(* IEC 61131-3 sources: SemaPLC/sema-plc-benchmark/spec2control-benchmark/data/st-baseline/waste_water_treatment_facility/pous/programs, 8 files *)

(* ---- main.st ---- *)
PROGRAM main
VAR
	Heartbeat : bool;
END_VAR

(* Entry point required by OpenPLC Editor v4. The process sections run as parallel program instances under task0; main only provides a scan heartbeat. *)
Heartbeat := NOT Heartbeat;

END_PROGRAM

(* ---- Section10.st ---- *)
PROGRAM Section10
VAR
	FT_901_FlowRate : real;
	LS_901_LevelPercent : real;
	P_901A_Running : bool;
	P_901B_Running : bool;
	P_901AB_DutyActiveIsA : bool;
	P_901AB_SwitchedDueToDuty : bool;
	P_901AB_SwitchedDueToFailure : bool;
	FT_901 : ANALOG_IN;
	LS_901 : ANALOG_IN;
	P_901A : MOTOR_ON_OFF;
	P_901B : MOTOR_ON_OFF;
	XV_102 : VALVE_ON_OFF;
	P_901AB : DUTY_STANDBY;
	DutyTimer_TON : TON;
	FailA_TON : TON;
	FailB_TON : TON;
	SwitchoverDelay_TON : TON;
	AnyRunning_OR : bool;
	StartBand_AND : bool;
	LevelAbove60_GT : bool;
	LevelAbove40_GT : bool;
	LevelAbove85_GT : bool;
	StartRequest_OR : bool;
	FlowLessThan15_GT : bool;
	FailCondA_AND : bool;
	FailCondB_AND : bool;
	Failure_OR : bool;
	StartCmdA_OR : bool;
	StartCmdB_OR : bool;
	PumpA_Inhibit_OR : bool;
	PumpB_Inhibit_OR : bool;
	BothPumpsFailed_AND : bool;
END_VAR

FT_901(
    Alarm_Enable := TRUE);
LS_901(
    PV_High := 90.0,
    Alarm_Enable := TRUE);
FlowLessThan15_GT := (REAL#15.0 > FT_901.PV);
FailCondA_AND := P_901A.FB_Running AND FlowLessThan15_GT;
FailA_TON(
    IN := FailCondA_AND,
    PT := T#10s);
PumpA_Inhibit_OR := LS_901.Low_Alarm OR FailA_TON.Q OR P_901A.FB_Trip;
LevelAbove85_GT := (LS_901.PV > REAL#85.0);
FailCondB_AND := P_901B.FB_Running AND FlowLessThan15_GT;
FailB_TON(
    IN := FailCondB_AND,
    PT := T#10s);
PumpB_Inhibit_OR := LS_901.Low_Alarm OR FailB_TON.Q OR P_901B.FB_Trip;
StartCmdB_OR := LevelAbove85_GT OR P_901AB.CmdPumpB;
P_901B(
    Start_Cmd := StartCmdB_OR,
    MinRunTime := T#30m,
    Inhibit := PumpB_Inhibit_OR);
AnyRunning_OR := P_901A.FB_Running OR P_901B.FB_Running;
DutyTimer_TON(
    IN := AnyRunning_OR,
    PT := T#48h);
LevelAbove60_GT := (LS_901.PV > REAL#60.0);
LevelAbove40_GT := (LS_901.PV > REAL#40.0);
StartBand_AND := AnyRunning_OR AND LevelAbove40_GT;
StartRequest_OR := LevelAbove60_GT OR StartBand_AND;
Failure_OR := FailA_TON.Q OR FailB_TON.Q;
SwitchoverDelay_TON(
    IN := Failure_OR,
    PT := T#5s);
P_901AB(
    Enable := TRUE,
    StartRequest := StartRequest_OR,
    AlternateEnable := TRUE,
    DutyElapsed := DutyTimer_TON.Q,
    SwitchoverDelayElapsed := SwitchoverDelay_TON.Q,
    PumpA_RunFB := P_901A.FB_Running,
    PumpB_RunFB := P_901B.FB_Running,
    PumpA_Fault := FailA_TON.Q,
    PumpB_Fault := FailB_TON.Q);
StartCmdA_OR := LevelAbove85_GT OR P_901AB.CmdPumpA;
P_901A(
    Start_Cmd := StartCmdA_OR,
    MinRunTime := T#30m,
    Inhibit := PumpA_Inhibit_OR);
BothPumpsFailed_AND := FailA_TON.Q AND FailB_TON.Q;
XV_102(
    Inhibit := BothPumpsFailed_AND);

(* Outputs published to other sections / HMI. *)
FT_901_FlowRate := FT_901.PV;
LS_901_LevelPercent := LS_901.PV;
P_901A_Running := P_901A.FB_Running;
P_901B_Running := P_901B.FB_Running;
P_901AB_DutyActiveIsA := P_901AB.ActiveIsA;
P_901AB_SwitchedDueToDuty := P_901AB.SwitchedDueToDuty;
P_901AB_SwitchedDueToFailure := P_901AB.SwitchedDueToFailure;

END_PROGRAM

(* ---- Section11.st ---- *)
PROGRAM Section11
VAR
	FIT_104_InfluentFlow_PV : real;
	FIC_106_SP_From_FFIC_107 : real;
	FIT_104 : ANALOG_IN;
	FFIC_107 : RATIO_CONTROL;
	FIC_106 : PID_BASIC;
	CD_1001 : MOTOR_VSD;
	PV_101 : VALVE_ELECTRIC;
	XV_102 : VALVE_ON_OFF;
	PumpInhibitAggregator : bool;
	RatioCtrlInhibitAggregator : bool;
	PumpOpenedInverter : bool;
END_VAR

FIT_104(
    Scaling_Slope := 6.25,
    Scaling_Offset := -25.0,
    Alarm_Enable := TRUE);
FIC_106(
    AUTO := TRUE,
    PV := CD_1001.FB_ActualSpeed,
    SP := FFIC_107.SlaveSP,
    MV_MIN := 0.0,
    MV_MAX := 100.0,
    Deviation_Limit := 3.0);
PV_101(
    Open_Limit := 100.0,
    Close_Limit := 0.0);
XV_102();
PumpOpenedInverter := NOT XV_102.FB_Opened;
PumpInhibitAggregator := PumpOpenedInverter OR FIT_104.Low_Alarm OR FIT_104.General_Fault OR XV_102.Alarm_General OR XV_102.Alarm_Position_Error OR PV_101.Alarm OR PV_101.Position_Error OR CD_1001.Alarm_Comm_Fail OR CD_1001.FB_Fault OR CD_1001.Alarm_Speed_Deviation;
CD_1001(
    Speed_SP := FIC_106.XOUT,
    Inhibit := PumpInhibitAggregator);
RatioCtrlInhibitAggregator := FIT_104.Low_Alarm OR FIT_104.High_Alarm OR FIT_104.General_Fault OR CD_1001.FB_Fault OR CD_1001.Alarm_Comm_Fail OR CD_1001.Alarm_Speed_Deviation;
FFIC_107(
    Auto := TRUE,
    PrimaryPV := FIT_104.PV,
    SecondaryPV := CD_1001.FB_ActualSpeed,
    RatioSP := 2.5,
    Bias := 0.0,
    MV_MIN := 0.0,
    MV_MAX := 100.0,
    Inhibit := RatioCtrlInhibitAggregator);

(* Outputs published to other sections / HMI. *)
FIT_104_InfluentFlow_PV := FIT_104.PV;
FIC_106_SP_From_FFIC_107 := FFIC_107.SlaveSP;

END_PROGRAM

(* ---- Section12.st ---- *)
PROGRAM Section12
VAR
	IIC101_Raw_mA : real;
	LV104_Raw_mA : real;
	IIC101_Solids_PV : real;
	IIC103_MV_to_PV102 : real;
	LV104_Level_PV : real;
	IIC_101 : ANALOG_IN;
	LV_104 : ANALOG_IN;
	IIC_103 : PID_BASIC;
	IIC_105 : BOOL_INPUT;
	PV_102 : VALVE_ELECTRIC;
	OC_1101 : VALVE_ON_OFF;
	OdorNotActive_NOT : bool;
	PIDInhibit_OR : bool;
	ValveInhibit_OR : bool;
END_VAR

IIC_101(
    Raw_Signal := IIC101_Raw_mA,
    Scaling_Slope := 0.625,
    Scaling_Offset := -2.5,
    Alarm_Enable := TRUE);
LV_104(
    Raw_Signal := LV104_Raw_mA,
    PV_High := 85.0,
    Scaling_Slope := 6.25,
    Scaling_Offset := -25.0,
    Alarm_Enable := TRUE);
PIDInhibit_OR := LV_104.High_Alarm OR IIC_101.General_Fault;
OC_1101(
    Timeout := T#10s);
IIC_105(
    Bool_In := OC_1101.FB_Opened);
OdorNotActive_NOT := NOT IIC_105.Bool_Out;
ValveInhibit_OR := OdorNotActive_NOT OR PV_102.Position_Error;
PV_102(
    Control_Signal := IIC_103.XOUT,
    Manual_Mode := FALSE,
    Open_Limit := 100.0,
    Close_Limit := 0.0,
    Timeout := T#30s,
    Inhibit := ValveInhibit_OR);
IIC_103(
    AUTO := TRUE,
    PV := IIC_101.PV,
    SP := 6.5,
    MV_MIN := 10.0,
    MV_MAX := 90.0,
    X0 := PV_102.Feedback_Pos,
    KP := 3.0,
    TR := 1.2,
    TD := 0.3,
    PV_High := 8.0,
    PV_Low := 4.0,
    Inhibit := PIDInhibit_OR);

(* Outputs published to other sections / HMI. *)
IIC101_Solids_PV := IIC_101.PV;
IIC103_MV_to_PV102 := IIC_103.XOUT;
LV104_Level_PV := LV_104.PV;

END_PROGRAM

(* ---- Section2.st ---- *)
PROGRAM Section2
VAR
	LS_101_WetWellLevel_PV_m : real;
	FT_101_InfluentFlow_PV_m3ph : real;
	PIC_101_WetWellLevel_MV_Pct : real;
	P_101A_Speed_Command_Pct : real;
	P_101B_Speed_Command_Pct : real;
	P101_LevelTrips_Active : bool;
	VG101_Inhibit_Active : bool;
	BS101_Disable_Active : bool;
	P_101A_Start_Cmd : bool;
	P_101B_Start_Cmd : bool;
	FT_101 : ANALOG_IN;
	LS_101 : ANALOG_IN;
	PIC_101 : PID_BASIC;
	P_101A : MOTOR_VSD;
	P_101B : MOTOR_VSD;
	XV_101 : VALVE_ON_OFF;
	BS_101 : BOOL_INPUT;
	VG_101 : MOTOR_ON_OFF;
	P101_LevelTrips_OR : bool;
	VG101_Inhibit_OR : bool;
	BS101_Disable_OR : bool;
	PID_Output_Positive_GT : bool;
	P101_LevelTrips_NOT : bool;
	PumpRunEnable_AND : bool;
	StartA_NOT : bool;
	StartB_NOT : bool;
	P101A_Running_NOT : bool;
	P101A_Failure_OR : bool;
	P101B_Start_AND : bool;
	LS101_HighAlarm_NOT : bool;
END_VAR

FT_101(
    Scaling_Slope := 31.25,
    Scaling_Offset := -125.0,
    Alarm_Enable := TRUE);
LS_101(
    PV_High := 8.5,
    PV_Low := 1.5,
    Scaling_Slope := 0.625,
    Scaling_Offset := -2.5,
    Alarm_Enable := TRUE);
PIC_101(
    AUTO := TRUE,
    PV := LS_101.PV,
    SP := 5.5,
    MV_MIN := 30.0,
    MV_MAX := 90.0,
    X0 := 0.0,
    KP := -2.0,
    TR := 1.5,
    TD := 0.3,
    Deviation_Limit := 0.1);
P101_LevelTrips_OR := PIC_101.PV_Low_Alarm OR PIC_101.PV_High_Alarm OR LS_101.High_Alarm;
P101_LevelTrips_NOT := NOT P101_LevelTrips_OR;
PumpRunEnable_AND := P101_LevelTrips_NOT;
StartA_NOT := NOT PumpRunEnable_AND;
P_101A(
    Start_Cmd := PumpRunEnable_AND,
    Stop_Cmd := StartA_NOT,
    Speed_SP := PIC_101.XOUT,
    Inhibit := P101_LevelTrips_OR);
P101A_Running_NOT := NOT P_101A.FB_Running;
P101A_Failure_OR := P_101A.FB_Fault OR P101A_Running_NOT;
P101B_Start_AND := PumpRunEnable_AND AND P101A_Failure_OR;
StartB_NOT := NOT P101B_Start_AND;
P_101B(
    Start_Cmd := P101B_Start_AND,
    Stop_Cmd := StartB_NOT,
    Speed_SP := PIC_101.XOUT,
    Inhibit := P101_LevelTrips_OR);
LS101_HighAlarm_NOT := NOT LS_101.High_Alarm;
XV_101(
    Open_Cmd := LS101_HighAlarm_NOT,
    Close_Cmd := LS_101.High_Alarm);
BS101_Disable_OR := PIC_101.PV_Low_Alarm OR LS_101.Low_Alarm;
BS_101(
    Bool_In := BS101_Disable_OR);
VG101_Inhibit_OR := LS_101.Low_Alarm OR FT_101.Low_Alarm;
VG_101(
    Inhibit := VG101_Inhibit_OR);
PID_Output_Positive_GT := (0.0 > 0.0);

(* Outputs published to other sections / HMI. *)
P101_LevelTrips_Active := P101_LevelTrips_OR;
VG101_Inhibit_Active := VG101_Inhibit_OR;
BS101_Disable_Active := BS101_Disable_OR;
P_101A_Start_Cmd := PumpRunEnable_AND;
P_101B_Start_Cmd := P101B_Start_AND;
LS_101_WetWellLevel_PV_m := LS_101.PV;
FT_101_InfluentFlow_PV_m3ph := FT_101.PV;
PIC_101_WetWellLevel_MV_Pct := PIC_101.XOUT;
P_101A_Speed_Command_Pct := P_101A.Speed_Out;
P_101B_Speed_Command_Pct := P_101B.Speed_Out;

END_PROGRAM

(* ---- Section4.st ---- *)
PROGRAM Section4
VAR
	FT301_InfluentFlow_PV : real;
	FT302_SludgeFlow_PV : real;
	LS301_WeirLevel_PV : real;
	PS301_SludgePressure_PV : real;
	FT302_SludgeFlow_SP : real;
	FT_301 : ANALOG_IN;
	FT_302 : ANALOG_IN;
	LS_301 : ANALOG_IN;
	PS_301 : ANALOG_IN;
	SS_301 : DIGITAL_IN;
	FV_102 : VALVE_ELECTRIC;
	FFIC_303 : RATIO_CONTROL;
	FIC_302 : PID_BASIC;
	FlowAboveCutoff_GT : bool;
	MasterInhibit_OR : bool;
END_VAR

FT_301(
    Alarm_Enable := TRUE);
FT_302(
    Alarm_Enable := TRUE);
LS_301(
    PV_High := 5.0,
    PV_Low := 2.0,
    Alarm_Enable := TRUE);
PS_301();
SS_301();
FlowAboveCutoff_GT := (FT_301.PV > 50.0);
MasterInhibit_OR := LS_301.High_Alarm OR LS_301.Low_Alarm OR FT_301.High_Alarm OR FT_301.Low_Alarm OR FT_301.General_Fault OR FT_302.High_Alarm OR FT_302.Low_Alarm OR FT_302.General_Fault OR FIC_302.Deviation_Alarm OR FV_102.Position_Error OR FV_102.Alarm OR SS_301.DI_Out;
FFIC_303(
    Auto := FlowAboveCutoff_GT,
    PrimaryPV := FT_301.PV,
    SecondaryPV := FT_302.PV,
    RatioSP := 0.3,
    Bias := 0.0,
    TrimKp := 0.0,
    TrimTi := T#0s,
    MV_MIN := 0.0,
    MV_MAX := 200.0,
    Inhibit := MasterInhibit_OR);
FIC_302(
    AUTO := FlowAboveCutoff_GT,
    PV := FT_302.PV,
    SP := FFIC_303.SlaveSP,
    MV_MIN := 0.0,
    MV_MAX := 100.0,
    Deviation_Limit := 10.0,
    Inhibit := MasterInhibit_OR);
FV_102(
    Control_Signal := FIC_302.XOUT,
    Manual_Mode := MasterInhibit_OR,
    Manual_Position := 0.0,
    Inhibit := MasterInhibit_OR);

(* Outputs published to other sections / HMI. *)
FT301_InfluentFlow_PV := FT_301.PV;
FT302_SludgeFlow_PV := FT_302.PV;
LS301_WeirLevel_PV := LS_301.PV;
PS301_SludgePressure_PV := PS_301.PV;
FT302_SludgeFlow_SP := FFIC_303.SlaveSP;

END_PROGRAM

(* ---- Section7.st ---- *)
PROGRAM Section7
VAR
	PT_601A_DischargePressure_PV : real;
	PT_601B_DischargePressure_PV : real;
	CL_601_ActiveIsA : bool;
	PS_601_ActiveIsA : bool;
	CL_601A : MOTOR_ON_OFF;
	CL_601B : MOTOR_ON_OFF;
	PS_601A : MOTOR_ON_OFF;
	PS_601B : MOTOR_ON_OFF;
	PT_601A : ANALOG_IN;
	PT_601B : ANALOG_IN;
	LS_601 : DIGITAL_IN;
	VS_601A : VALVE_ELECTRIC;
	VS_601B : VALVE_ELECTRIC;
	CL_601A_CL_601B : DUTY_STANDBY;
	PS_601A_PS_601B : DUTY_STANDBY;
	Clar_MinRunTimer_TON : TON;
	Clar_DutyTimer_TON : TON;
	Clar_SwitchoverDelay_TON : TON;
	Pump_MinRunTimer_TON : TON;
	Pump_DutyTimer_TON : TON;
	Pump_SwitchoverDelay_TON : TON;
	ClarifierAnyRunning_OR : bool;
	ClarifierNoneRunning_NOT : bool;
	PumpAnyRunning_OR : bool;
	PumpNoneRunning_NOT : bool;
	PS601A_Inhibit_OR : bool;
	PS601B_Inhibit_OR : bool;
END_VAR

LS_601();
CL_601B(
    Start_Cmd := CL_601A_CL_601B.CmdPumpB,
    Start_Delay := T#5s,
    MinRunTime := T#30m,
    Inhibit := LS_601.DI_Out);
ClarifierAnyRunning_OR := CL_601A.FB_Running OR CL_601B.FB_Running;
Clar_DutyTimer_TON(
    IN := ClarifierAnyRunning_OR,
    PT := T#72h);
Clar_MinRunTimer_TON(
    IN := ClarifierAnyRunning_OR,
    PT := T#30m);
ClarifierNoneRunning_NOT := NOT ClarifierAnyRunning_OR;
Clar_SwitchoverDelay_TON(
    IN := ClarifierNoneRunning_NOT,
    PT := T#10s);
CL_601A_CL_601B(
    Enable := TRUE,
    StartRequest := TRUE,
    AlternateEnable := TRUE,
    DutyElapsed := Clar_DutyTimer_TON.Q,
    MinRunElapsed := Clar_MinRunTimer_TON.Q,
    SwitchoverDelayElapsed := Clar_SwitchoverDelay_TON.Q,
    PumpA_RunFB := CL_601A.FB_Running,
    PumpB_RunFB := CL_601B.FB_Running,
    PumpA_Fault := CL_601A.FB_Trip,
    PumpB_Fault := CL_601B.FB_Trip,
    Inhibit := LS_601.DI_Out);
CL_601A(
    Start_Cmd := CL_601A_CL_601B.CmdPumpA,
    Start_Delay := T#5s,
    MinRunTime := T#30m,
    Inhibit := LS_601.DI_Out);
PT_601A(
    PV_Low := 25.0,
    Alarm_Enable := TRUE);
PS601A_Inhibit_OR := PT_601A.Low_Alarm OR LS_601.DI_Out;
PT_601B(
    PV_Low := 25.0,
    Alarm_Enable := TRUE);
PS601B_Inhibit_OR := PT_601B.Low_Alarm OR LS_601.DI_Out;
PS_601B(
    Start_Cmd := PS_601A_PS_601B.CmdPumpB,
    Start_Delay := T#5s,
    MinRunTime := T#30m,
    Inhibit := PS601B_Inhibit_OR);
PumpAnyRunning_OR := PS_601A.FB_Running OR PS_601B.FB_Running;
Pump_DutyTimer_TON(
    IN := PumpAnyRunning_OR,
    PT := T#72h);
Pump_MinRunTimer_TON(
    IN := PumpAnyRunning_OR,
    PT := T#30m);
PumpNoneRunning_NOT := NOT PumpAnyRunning_OR;
Pump_SwitchoverDelay_TON(
    IN := PumpNoneRunning_NOT,
    PT := T#10s);
PS_601A_PS_601B(
    Enable := TRUE,
    StartRequest := TRUE,
    AlternateEnable := TRUE,
    DutyElapsed := Pump_DutyTimer_TON.Q,
    MinRunElapsed := Pump_MinRunTimer_TON.Q,
    SwitchoverDelayElapsed := Pump_SwitchoverDelay_TON.Q,
    PumpA_RunFB := PS_601A.FB_Running,
    PumpB_RunFB := PS_601B.FB_Running,
    PumpA_Fault := PS_601A.FB_Trip,
    PumpB_Fault := PS_601B.FB_Trip,
    Inhibit := LS_601.DI_Out);
PS_601A(
    Start_Cmd := PS_601A_PS_601B.CmdPumpA,
    Start_Delay := T#5s,
    MinRunTime := T#30m,
    Inhibit := PS601A_Inhibit_OR);
VS_601A(
    Open_Limit := 100.0,
    Close_Limit := 0.0);
VS_601B(
    Open_Limit := 100.0,
    Close_Limit := 0.0);

(* Outputs published to other sections / HMI. *)
PT_601A_DischargePressure_PV := PT_601A.PV;
PT_601B_DischargePressure_PV := PT_601B.PV;
CL_601_ActiveIsA := CL_601A_CL_601B.ActiveIsA;
PS_601_ActiveIsA := PS_601A_PS_601B.ActiveIsA;

END_PROGRAM

(* ---- Section9.st ---- *)
PROGRAM Section9
VAR
	FT_801_EffluentFlow_PV : real;
	CL_801_ChlorineFlow_SP : real;
	DC_801_DechlorFlow_SP : real;
	XV_106_FullyOpen_FB : bool;
	CL_801_Running_FB : bool;
	DC_801_Running_FB : bool;
	FT_801 : ANALOG_IN;
	FIC_101 : RATIO_CONTROL;
	FIC_102 : RATIO_CONTROL;
	CL_801 : MOTOR_VSD;
	DC_801 : MOTOR_VSD;
	LV_105 : VALVE_ELECTRIC;
	XV_106 : VALVE_ON_OFF;
	UV_801 : MOTOR_ON_OFF;
	CL_RatioMinCalc : real;
	CL_RatioMaxCalc : real;
	DC_RatioMinCalc : real;
	DC_RatioMaxCalc : real;
	ValveNotOpen : bool;
	CL_NotRunning : bool;
	ChemActive : bool;
	LV_105_AnyAlarm : bool;
	XV_106_AnyAlarm : bool;
	CL_801_Inh_OR1 : bool;
	CL_801_Inh_OR2 : bool;
	CL_801_Inh_OR3 : bool;
	DC_801_Inh_OR1 : bool;
	DC_801_Inh_OR2 : bool;
	FT_801_AnyFault_OR1 : bool;
	FT_801_AnyFault_OR2 : bool;
	FIC_102_Inh_OR1 : bool;
END_VAR

FT_801(
    Scaling_Slope := 62.5,
    Scaling_Offset := -250.0,
    Alarm_Enable := TRUE);
XV_106(
    Timeout := T#5s);
ValveNotOpen := NOT XV_106.FB_Opened;
CL_801_Inh_OR1 := ValveNotOpen OR FT_801.Low_Alarm;
XV_106_AnyAlarm := XV_106.Alarm_Position_Error OR XV_106.Alarm_General;
CL_801_Inh_OR2 := CL_801_Inh_OR1 OR XV_106_AnyAlarm;
LV_105(
    Timeout := T#5s);
LV_105_AnyAlarm := LV_105.Position_Error OR LV_105.Alarm;
CL_801_Inh_OR3 := CL_801_Inh_OR2 OR LV_105_AnyAlarm;
CL_801(
    Speed_SP := FIC_101.SlaveSP,
    Inhibit := CL_801_Inh_OR3);
CL_RatioMaxCalc := FT_801.PV * 3.0;
CL_RatioMinCalc := FT_801.PV * 2.0;
FT_801_AnyFault_OR1 := FT_801.Low_Alarm OR FT_801.High_Alarm;
FT_801_AnyFault_OR2 := FT_801_AnyFault_OR1 OR FT_801.General_Fault;
FIC_101(
    Auto := TRUE,
    PrimaryPV := FT_801.PV,
    SecondaryPV := CL_801.FB_ActualSpeed,
    RatioSP := 2.5,
    MV_MIN := CL_RatioMinCalc,
    MV_MAX := CL_RatioMaxCalc,
    Inhibit := FT_801_AnyFault_OR2);
CL_NotRunning := NOT CL_801.FB_Running;
DC_801_Inh_OR1 := LV_105_AnyAlarm OR FT_801.Low_Alarm;
DC_801_Inh_OR2 := DC_801_Inh_OR1 OR CL_NotRunning;
DC_801(
    Speed_SP := FIC_102.SlaveSP,
    Inhibit := DC_801_Inh_OR2);
DC_RatioMaxCalc := FT_801.PV * 1.5;
DC_RatioMinCalc := FT_801.PV * 1.0;
FIC_102_Inh_OR1 := FT_801_AnyFault_OR2 OR CL_NotRunning;
FIC_102(
    Auto := TRUE,
    PrimaryPV := FT_801.PV,
    SecondaryPV := DC_801.FB_ActualSpeed,
    RatioSP := 1.2,
    MV_MIN := DC_RatioMinCalc,
    MV_MAX := DC_RatioMaxCalc,
    Inhibit := FIC_102_Inh_OR1);
ChemActive := CL_801.FB_Running OR DC_801.FB_Running;
UV_801(
    Inhibit := ChemActive);

(* Outputs published to other sections / HMI. *)
FT_801_EffluentFlow_PV := FT_801.PV;
CL_801_ChlorineFlow_SP := FIC_101.SlaveSP;
DC_801_DechlorFlow_SP := FIC_102.SlaveSP;
XV_106_FullyOpen_FB := XV_106.FB_Opened;
CL_801_Running_FB := CL_801.FB_Running;
DC_801_Running_FB := DC_801.FB_Running;

END_PROGRAM
